(* PLC project v0.5.4_.project, CODESYS CODESYS V3.5 SP19 Patch 1 *)
(* stored: creationDateTime 2026-08-03T23:41:10.3091042, modificationDateTime 2026-08-03T23:40:10.7089817 *)

PROGRAM PRG_01_Inputs_LD
  VAR_OUTPUT
    PowerContactorEngaged : BOOL;
    M1BrakeFeedback : BOOL;
  END_VAR
  VAR
    instPowerContactorEngaged : FB_Input;
    instM1BrakeFeedback : FB_Input;
  END_VAR

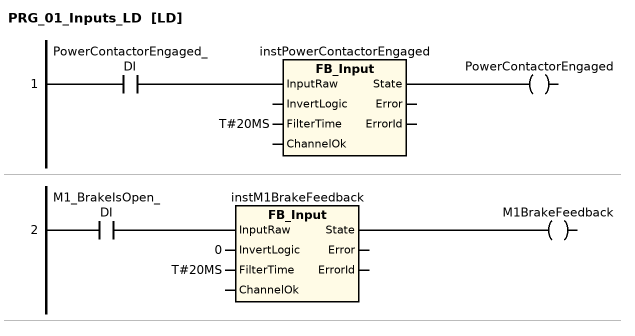
(* LD diagram, written out as Structured Text *)

instPowerContactorEngaged(InputRaw := PowerContactorEngaged_DI, InvertLogic := , FilterTime := T#20MS, ChannelOk := );
PowerContactorEngaged := instPowerContactorEngaged.State;

instM1BrakeFeedback(InputRaw := M1_BrakeIsOpen_DI, InvertLogic := 0, FilterTime := T#20MS, ChannelOk := );
M1BrakeFeedback := instM1BrakeFeedback.State;
END_PROGRAM
